(* IEC 61131-3 sources: llm-plc-st-eval/data/processed_v2/gpt-4o/B6/zero_shot, 3 files *)

(* ---- ejec_1.st ---- *)
FUNCTION_BLOCK FB_Baliza
VAR
    alarma : BOOL; // Variable de entrada: indica si la alarma está activa
    lampara : BOOL; // Variable de salida: controla el estado de la lámpara
    ton : TON; // Temporizador TON para controlar el parpadeo
    estado_parpadeo : BOOL; // Estado interno para el parpadeo
END_VAR

// Inicialización del temporizador
ton(IN := estado_parpadeo, PT := T#1S);

// Lógica de control de la baliza
IF alarma THEN
    // Si la alarma está activa, alternar el estado de parpadeo
    IF ton.Q THEN
        estado_parpadeo := NOT estado_parpadeo; // Cambiar el estado de parpadeo
        ton(IN := FALSE); // Reiniciar el temporizador
    ELSE
        ton(IN := TRUE); // Activar el temporizador
    END_IF;
    lampara := estado_parpadeo; // Actualizar el estado de la lámpara
ELSE
    // Si no hay alarma, la lámpara está apagada
    lampara := FALSE;
    estado_parpadeo := FALSE; // Reiniciar el estado de parpadeo
    ton(IN := FALSE); // Asegurarse de que el temporizador esté desactivado
END_IF;
END_FUNCTION_BLOCK

(* ---- ejec_2.st ---- *)
FUNCTION_BLOCK FB_Baliza
VAR_INPUT
    alarma : BOOL; // Variable de entrada que indica si hay una condición de alarma
END_VAR

VAR_OUTPUT
    lampara : BOOL; // Variable de salida que controla el estado de la lámpara
END_VAR

VAR
    ton : TON; // Temporizador para controlar el parpadeo
    estado : BOOL; // Estado interno para alternar el parpadeo
END_VAR

// Inicialización del temporizador
ton(IN := estado, PT := T#1S);

// Lógica de control de la baliza
IF alarma THEN
    // Si la alarma está activa, alternar el estado de la lámpara
    IF ton.Q THEN
        estado := NOT estado; // Cambiar el estado interno
        ton(IN := FALSE); // Reiniciar el temporizador
    ELSE
        ton(IN := TRUE); // Activar el temporizador
    END_IF;
    lampara := estado; // Actualizar el estado de la lámpara
ELSE
    // Si no hay alarma, la lámpara permanece apagada
    lampara := FALSE;
    estado := FALSE; // Reiniciar el estado interno
    ton(IN := FALSE); // Asegurarse de que el temporizador esté apagado
END_IF;

END_FUNCTION_BLOCK

(* ---- ejec_3.st ---- *)
FUNCTION_BLOCK FB_Baliza
VAR_INPUT
    alarma : BOOL; // Variable de entrada que indica si la alarma está activa
END_VAR

VAR_OUTPUT
    lampara : BOOL; // Variable de salida que controla el estado de la lámpara
END_VAR

VAR
    timerBlink : TON; // Temporizador para controlar el parpadeo
    estadoParpadeo : BOOL; // Estado interno para alternar el parpadeo
END_VAR

// Inicialización del temporizador
timerBlink(IN := estadoParpadeo, PT := T#1S);

IF alarma THEN
    // Si la alarma está activa, controlar el parpadeo
    IF timerBlink.Q THEN
        estadoParpadeo := NOT estadoParpadeo; // Alternar el estado de parpadeo
        timerBlink(IN := estadoParpadeo); // Reiniciar el temporizador
    END_IF;
    lampara := estadoParpadeo; // Actualizar la salida de la lámpara
ELSE
    // Si no hay alarma, la lámpara permanece apagada
    lampara := FALSE;
    estadoParpadeo := FALSE; // Reiniciar el estado de parpadeo
    timerBlink(IN := FALSE); // Asegurarse de que el temporizador esté detenido
END_IF;

END_FUNCTION_BLOCK
